// TIA Portal V21 export
// export: Created 2026-11-21T11:47:44.3576274Z, ExportSetting WithDefaults, DisplayName Totally Integrated Automation Portal, DisplayVersion V21, DisplayName STEP 7 Professional, DisplayVersion V21, DisplayName STEP 7 Safety, DisplayVersion V21, DisplayName Tech WebApplication, DisplayVersion V21, DisplayName WinCC Basic/Comfort/Advanced, DisplayVersion V21, DisplayName WinCC Unified, DisplayVersion V21
FUNCTION_BLOCK "Mixed"   // FB12, LAD
TITLE = Mixed languages
{ S7_Optimized_Access := 'TRUE' }
VERSION : 0.1
// A ladder block with an SCL and an STL network.
// stored: AutoNumber true, IsIECCheckEnabled false, IsRetainMemResEnabled false, MemoryReserve 100, SetENOAutomatically false, UDAEnableTagReadback false
   VAR_INPUT
      start : Bool;
      stop : Bool;
      door : Bool;
   END_VAR
   VAR_OUTPUT
      motor : Bool;
      lamp : Bool;
      fault : Bool;
   END_VAR
   VAR
      latched : Bool;
      edgeMemory : Bool;
   END_VAR
BEGIN

REGION Network 1: Ladder
   // A ladder network first.
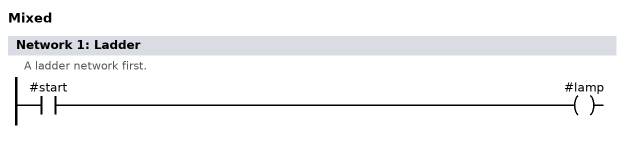
   RUNG wire#powerrail
      Contact( #start )
      Coil( #lamp )
   END_RUNG
   // the same network as SCL:
   #lamp := #start;
END_REGION

REGION Network 2 (SCL): Structured text
   // An SCL network inside a ladder block.
   #motor := #start AND NOT #stop;
END_REGION

NETWORK
TITLE = Statement list
// An STL network inside a ladder block.
      A     #door;
      AN    #stop;
      =     #fault;
END_FUNCTION_BLOCK
